FUNCTION_BLOCK fb_Dev_ControlValve_Modulating EXTENDS abs_fb_Device
VAR_INPUT
	inpValvePosition	: LREAL;
END_VAR

VAR
	transMantoAuto	: R_TRIG;
	transAutoToMan	: F_TRIG;
END_VAR

VAR PERSISTENT
	HMI				: ST_ControlValve_Modulating_HMI_Interface;
	_valvePosition	: LREAL;
END_VAR


VAR_OUTPUT
	outValvePosition	: LREAL;
	stsValveFeedback	: LREAL;
END_VAR

DeviceLogic();
Interlock.name := _DeviceName;
Interlock(inpConfig := _dataInterlock);

faultHandler();

transManToAuto(CLK:=_inAuto);
transAutoToMan(CLK:=_inAuto);

stsValveFeedback := inpValvePosition;

// Maintain valve position during man/auto machine state changes
IF transManToAuto.Q THEN
	_valvePosition := HMI.ocmdValvePosition;
END_IF

IF transAutoToMan.Q THEN
	HMI.ocmdValvePosition := _valvePosition;
END_IF

IF NOT stsFaulted AND Interlock.outInterlockOK THEN
	IF _inAuto THEN
		outValvePosition := _valvePosition;
	ELSE
		outValvePosition := HMI.ocmdValvePosition;
	END_IF
END_IF

HMI.stsValveFeedback := stsValveFeedback;
HMI.stsValvePosition := outValvePosition;
HMI.HMIbaseDevice := HMIBaseDevice;

METHOD faultHandler : BOOL
VAR_INPUT
END_VAR
IF stsValveFeedback < -1 AND _warnChannels[1] = '' THEN
	sendWarning('Valve feedback not present', 1);
END_IF
END_METHOD

PROPERTY valvePosition : LREAL
GET
valvePosition := _valvePosition;
END_GET
SET
_valvePosition := valvePosition;
END_SET
END_PROPERTY

END_FUNCTION_BLOCK

(* stored: Version 1.1.0.1
   POU fb_Dev_ControlValve_Modulating: Id {89888e0f-f91a-4412-8354-ec910db7043f}, SpecialFunc None
   Method faultHandler: Id {adf71b67-ffd5-4f27-bbed-e6c2244bc31f}
   Property valvePosition: Id {fd4b2016-bcc6-4cab-895b-90d88535bd1f}
   Get Get: Id {b82cfbac-57a6-4808-bcff-8cb24271bbb6}
   Set Set: Id {802320db-e8e9-4dc2-bba0-e1b6ceff50e0} *)
